(* IEC 61131-3 sources: Lasal-MCP/examples/SampleSource/2_PumpControlSolution/Stations/MachineControl/MachineControl/Class/SafetyCDIAS_Base (part 2) *)

        p_HandlePDOWrite^$USINT := VARAN_DO_NO_RUN;
      end_if;

      ud_LocalMoveDestAddr := pPDOWriteData$UDINT;
    end_if;

    if sd_VaranType = 1 then

      //add data object for TDO write
      sd_retval := MasterConnect.AddWrDO( ud_dol_type   := VARAN_DOL_ISO
                                        , p_ud_handle	  := ( #p_HandleTDOWrite )$^UDINT
                                        , ud_address	  := ui_MyPlace + OFFSET_STDO_DATA
                                        , ud_length	    := STDO_LENGTH
                                        , p_ud_data	    := ( #p_us_Handle_TDO_Write )$^UDINT
                                        , ud_type			  := 1
                                        );

      //look for an error
      if ( sd_retval <> 0 ) then
        State.uiIO_Flags				          := 0;
        State.uiIO_Flags.NoCalibration	  := 1;
        State.uiIO_Flags.PhysicAccessOff  := 1;
        return;
      end_if;
    else  // for mover we have to say it's a single execution

      //add data object for TDO write
      sd_retval := MasterConnect.AddWrDO( ud_dol_type   := VARAN_DOL_ISO
                                        , p_ud_handle	  := ( #p_HandleTDOWrite )$^UDINT
                                        , ud_address	  := ui_MyPlace + OFFSET_STDO_DATA
                                        , ud_length	    := STDO_LENGTH
                                        , p_ud_data	    := ( #p_us_Handle_TDO_Write )$^UDINT
                                        , ud_type			  := 1 OR VM_SINGLE_ID
                                        );

      //look for an error
      if ( sd_retval <> 0 ) then
        State.uiIO_Flags				          := 0;
        State.uiIO_Flags.NoCalibration	  := 1;
        State.uiIO_Flags.PhysicAccessOff  := 1;
        return;
      end_if;

      (p_HandleTDOWrite$^USINT )^ := VARAN_DO_NO_RUN;
    end_if;

    // only for modules with outputs
    if Kennung <> CSDI16x_ID then

      //add data object for unsafe output write
      sd_retval := MasterConnect.AddWrDO( ud_dol_type   := VARAN_DOL_ISO
                                        , p_ud_handle	  := ( #p_HandleUnsafeOutWrite )$^UDINT
                                        , ud_address	  := ui_MyPlace + OFFSET_UNSAFE_VAR
                                        , ud_length	    := UNSAFE_OUT_LENGTH
                                        , p_ud_data	    := ( #p_ui_UnsafeOutWrite )$^UDINT
                                        , ud_type			  := 1
                                        );

      //look for an error
      if ( sd_retval <> 0 ) then
        State.uiIO_Flags				          := 0;
        State.uiIO_Flags.NoCalibration	  := 1;
        State.uiIO_Flags.PhysicAccessOff  := 1;
        return;
      end_if;
    end_if;

    //data object for LEDs, SSDO State, STDO State, SPDO DataLength and time sync handshake
    sd_retval := MasterConnect.AddRdDO( ud_dol_type   := VARAN_DOL_ISO
                                      , p_ud_handle   := ( #p_HandleLED )$^UDINT
                                      , ud_address    := ui_MyPlace + OFFSET_LED
                                      , ud_length     := 15
                                      , p_ud_data     := ( #p_ud_Handle_LED )$^UDINT
                                      , ud_type       := 1
                                      );

    //look for an error
    if ( sd_retval <> 0 ) then
      State.uiIO_Flags				          := 0;
      State.uiIO_Flags.NoCalibration	  := 1;
      State.uiIO_Flags.PhysicAccessOff  := 1;
      return;
    end_if;

    p_us_Handle_TDO_Read_Length   := p_ud_Handle_LED + (OFFSET_STDO_STATUS - OFFSET_LED);
    p_us_Handle_TDO_Read_Length^  := 0;

    pPDOReadLengthData := p_ud_Handle_LED + (OFFSET_SPDO_LENGTH - OFFSET_LED);
    pPDOReadLengthData^ := 0;

    p_us_Handle_TDO_Status_Write  := p_ud_Handle_LED + (OFFSET_STDO_STATUS_WRITE - OFFSET_LED);
    p_us_Handle_TDO_Status_Write^ := 0;

    p_us_Handle_TimeSyncHS_Read   := p_ud_Handle_LED + (OFFSET_TIMESYNC_HANDSHAKE - OFFSET_LED);
    p_us_Handle_TimeSyncHS_Read^  := 0;

    if sd_VaranType = 1 then

      //add data object for time sync handshake
      sd_retval := MasterConnect.AddWrDO( ud_dol_type   := VARAN_DOL_ISO
                                        , p_ud_handle	  := ( #p_Handle_TimeSyncHS_Write )$^UDINT
                                        , ud_address	  := ui_MyPlace + OFFSET_TIMESYNC_HANDSHAKE
                                        , ud_length	    := 1
                                        , p_ud_data	    := ( #p_us_Handle_TimeSyncHS_Write )$^UDINT
                                        , ud_type			  := 1
                                        );

    else  // for mover we have to say it's a single execution

      //add data object for TDO write
      sd_retval := MasterConnect.AddWrDO( ud_dol_type   := VARAN_DOL_ISO
                                        , p_ud_handle	  := ( #p_Handle_TimeSyncHS_Write )$^UDINT
                                        , ud_address	  := ui_MyPlace + OFFSET_TIMESYNC_HANDSHAKE
                                        , ud_length	    := 1
                                        , p_ud_data	    := ( #p_us_Handle_TimeSyncHS_Write )$^UDINT
                                        , ud_type			  := 1 OR VM_SINGLE_ID
                                        );
      (p_Handle_TimeSyncHS_Write$^USINT )^ := VARAN_DO_NO_RUN;
    end_if;

    //look for an error
    if ( sd_retval <> 0 ) then
      State.uiIO_Flags				          := 0;
      State.uiIO_Flags.NoCalibration	  := 1;
      State.uiIO_Flags.PhysicAccessOff  := 1;
      return;
    end_if;

    //add data object for TDO read
    sd_retval := MasterConnect.AddRdDO( ud_dol_type   := VARAN_DOL_ISO
                                      , p_ud_handle	  := ( #p_HandleTDORead )$^UDINT
                                      , ud_address	  := ui_MyPlace + OFFSET_STDO_DATA
                                      , ud_length	    := STDO_LENGTH
                                      , p_ud_data	    := ( #p_us_Handle_TDO_Read )$^UDINT
                                      , ud_type			  := 1
                                      );

    //look for an error
    if ( sd_retval <> 0 ) then
      State.uiIO_Flags				          := 0;
      State.uiIO_Flags.NoCalibration	  := 1;
      State.uiIO_Flags.PhysicAccessOff  := 1;
      return;
    end_if;

    // fast unsafe variables (only if activated)
    if ActivateFastUnsafeIOs then
      //add data object for fast unsafe output and input variables
      sd_retval :=  MasterConnect.AddRdWrDO(ud_dol_type       := VARAN_DOL_ISO
                                          , p_ud_handle       := ( #p_HandleFastUnsafeIOs )$^UDINT
                                          , ud_address_read   := ui_MyPlace + OFFSET_FAST_UNSAFE_IOS
                                          , ud_length_read    := 1
                                          , p_ud_data_read    := ( #p_us_Handle_FastUnsafeOutputs )$^UDINT
                                          , ud_address_write  := ui_MyPlace + OFFSET_FAST_UNSAFE_IOS
                                          , ud_length_write   := 1
                                          , p_ud_data_write   := ( #p_us_Handle_FastUnsafeInputs )$^UDINT
                                          , ud_type           := 1
                                          );

      //look for an error
      if ( sd_retval <> 0 ) then
        State.uiIO_Flags				          := 0;
        State.uiIO_Flags.NoCalibration	  := 1;
        State.uiIO_Flags.PhysicAccessOff  := 1;
        return;
      end_if;
    end_if;
  end_if;

END_FUNCTION

FUNCTION VIRTUAL SafetyCDIAS_Base::GetPointer2PDOBuffer
	VAR_OUTPUT
		ud_PDOBuffer 	: UDINT;
	END_VAR

  PDOOutputIsUsed := TRUE;

  //set pointer to address of buffer pointer
  ud_PDOBuffer := ( #PDOOutputBuffer )$UDINT;

END_FUNCTION

FUNCTION VIRTUAL SafetyCDIAS_Base::AddRoutingElement
	VAR_INPUT
		ud_SafeNumber 	: HDINT;
		ud_thisp 	      : UDINT;
		pObject 	      : ^PathInfoType;
	END_VAR
	VAR_OUTPUT
		sd_retval 	    : DINT;
	END_VAR
  VAR
  	p_RoutElement   : ^RoutElement;
    ui_PathLength   : UINT;
    NewElement      : BOOL;
  END_VAR

  if ( ( ud_SafeNumber <> 0 ) & ( ud_thisp <> NIL ) ) then
    if ui_CntRoutElements < MAX_NUMBER_ROUT_ELEMENTS then

      NewElement := TRUE;

      if ui_CntRoutElements then
        //check if object this-pointer already exists in routing table
        p_RoutElement := GetRoutingElementByThis( ud_thisp := ud_thisp );
      else
        p_RoutElement := NIL;
      end_if;

      if p_RoutElement = NIL then
        //add new element

        //set pointer to empty element on last position
        p_RoutElement := p_RoutTable + ( ui_CntRoutElements ) * sizeof(RoutElement);
      else
        // we don't have a new element, we just update an existing
        NewElement := FALSE;
      end_if;

      //add path

      // path isn't stored if it's the routing table of safe input module, because
      // it doesn't need the information
      if pObject^.p_us_Path & pObject^.p_us_PathComp
         & ((NewElement = TRUE) | ((NewElement = FALSE) & (p_RoutElement^.p_CompressedPath = NIL) & (p_RoutElement^.ui_ComprPathLen = 0))) // only if it isn't already set
         then

        // the whole object path isn't stored, because the path can't be used for routing of SDOs;
        // The length of the path varies and it's possible, that the path is too long
        // to transfer it in SDO header. Instead of it the compressed path is used for addressing.

        ui_PathLength := pObject^.ui_PathCompLen;
        p_RoutElement^.p_CompressedPath$pVoid := To_StdLib.Malloc(size := ui_PathLength);

        if ( p_RoutElement^.p_CompressedPath = NIL ) then

          State.uiIO_Flags                  := 0;
          State.uiIO_Flags.PhysicAccessOff 	:= 1;
          sd_retval                         :=-1;
          ClassState := _MemAllocFailed;
          return;

        end_if;

        // store compressed path into actual routing element
        To_StdLib.MemCpy(dest := p_RoutElement^.p_CompressedPath, source := pObject^.p_us_PathComp, size := ui_PathLength);
        p_RoutElement^.ui_ComprPathLen := ui_PathLength;
      elsif NewElement then

        // not routing table of safety CPU of safety output
        p_RoutElement^.p_CompressedPath := NIL;
        p_RoutElement^.ui_ComprPathLen  := 0;
      end_if;

      //insert data
      p_RoutElement^.ud_SafeNumber      := ud_SafeNumber;
      p_RoutElement^.ud_thisp           := ud_thisp;

      if NewElement then
        //increase counter
        ui_CntRoutElements += 1;
      end_if;

      sd_retval := 0;
    else

      sd_retval := -1;
      LogError("@ZZZZ (SafetyCDIAS_Base::AddRoutingElement) Maximum number of possible routing elements reached");
    end_if;
  else

    sd_retval := -1;

    if ud_SafeNumber = 0 then
      LogError("@ZZZZ (SafetyCDIAS_Base::AddRoutingElement) 0 is an invalid safety number");
    else
      LogError("@ZZZZ (SafetyCDIAS_Base::AddRoutingElement) NIL pointer given as this pointer");
    end_if;
  end_if;

END_FUNCTION

FUNCTION VIRTUAL SafetyCDIAS_Base::GetRoutingPointerByNumber
	VAR_INPUT
		ud_SafeNumber 	: HDINT;
	END_VAR
	VAR_OUTPUT
		ud_thisp 	      : UDINT;
	END_VAR
  VAR
  	i               : UINT;
    p_RoutElement   : ^RoutElement;
  END_VAR

  ud_thisp := 0;

  //no valid safety number
  if ( ud_SafeNumber = 0 ) then
    return;
  end_if;

  //set pointer on first routing element
  p_RoutElement := p_RoutTable;

  //check each element
  if ( ui_CntRoutElements > 0 ) then
    for i := 0 to ui_CntRoutElements - 1 by 1 do

      //if searched safety number is found, this-pointer is returned
      if ( p_RoutElement^.ud_SafeNumber = ud_SafeNumber ) then

        ud_thisp := p_RoutElement^.ud_thisp;
        return;

      end_if;

      //set pointer to next element
      p_RoutElement += sizeof ( RoutElement );

    end_for;
  end_if;

END_FUNCTION

FUNCTION VIRTUAL SafetyCDIAS_Base::GetRoutingPointerByPath
	VAR_INPUT
		p_ActObjectPath 	: ^USINT;
		ActPathLen 	      : UINT;
	END_VAR
	VAR_OUTPUT
		ud_thisp          : UDINT;
	END_VAR
  VAR
  	i                 : UINT;
    p_RoutElement     : ^RoutElement;
    retcode           : UINT;
  END_VAR

  ud_thisp := 0;

  //set pointer on first routing element
  p_RoutElement := p_RoutTable;

  //check each element
  if ( ui_CntRoutElements > 0 ) then
    for i := 0 to ui_CntRoutElements - 1 by 1 do

      if p_RoutElement^.p_CompressedPath & (p_RoutElement^.ui_ComprPathLen = ActPathLen) then

        //if searched path is found, this-pointer is returned
        retcode := To_StdLib.MemCmp(dest:= p_ActObjectPath, source:= p_RoutElement^.p_CompressedPath , size:= ActPathLen);

        if retcode = 0 then

          ud_thisp := p_RoutElement^.ud_thisp;
          return;

        end_if;
      end_if;

      //set pointer to next element
      p_RoutElement += sizeof ( RoutElement );

    end_for;
  end_if;

END_FUNCTION

FUNCTION VIRTUAL SafetyCDIAS_Base::ConfigSafetyInput
	VAR_INPUT
		ud_SafeNrCPU 	        : HDINT;
		ud_thisp 	            : UDINT;
		p_PDOBuffer 	        : ^UDINT;
		pMoveActive 	        : ^PDOMoveState;
		p_ud_HandleSourceDO 	: ^UDINT;
		p_ud_MoveSourceAddr 	: ^UDINT;
		p_ud_MoveSourceOffset : ^UDINT;
	END_VAR
	VAR_OUTPUT
		ud_SafeNrModul 	      : HDINT;
	END_VAR
  VAR
  	TempPathInfo          : PathInfoType;
  END_VAR

  ud_SafeNrModul := 0;

  if (State.uiIO_Flags = 0) then
    if ( ud_SafeNrCPU ) then

      // if pMoveActive is available, the data are sent to a CPU via VARAN => moving is possible
      if pMoveActive then
        // if input module is also accessed via VARAN => activate moving
        if b_VaranAvailable & (b_SafetyOnLocalCDIAS = FALSE) then
          // pdos are moved from csdi to cscp
          b_MoveCommandOutputActive := _Active;

          p_ud_MoveSourceAddr^      := pPDOReadData$UDINT;

          // Return DO Handle and Offset, Needed for Payload Move DOs
          if sd_VaranType = 1 then  // Return DO Handle
            p_ud_HandleSourceDO^    := p_HandlePDORead$UDINT;
          else                      // Return VaranDataMoversDO Handle
            p_ud_HandleSourceDO^    := 0;
          end_if;

          p_ud_MoveSourceOffset^    := 0;

          // Return DO Handle and Offset, Needed for Payload Move DOs
          if sd_VaranType = 1 then  // Return DO Handle
            p_ud_HandleSourceDO^    := p_HandlePDORead$UDINT;
          else                      // Return VaranDataMoversDO Handle
            p_ud_HandleSourceDO^    := ud_HandlePDOReadMoverDO;
          end_if;

          p_ud_MoveSourceOffset^    := 0;
        else
          // pdos are not moved from csdi to cscp or cscp to csto
          pMoveActive^              := _Inactive;
          b_MoveCommandOutputActive := _Inactive;
        end_if;
      else
        b_MoveCommandOutputActive   := _Inactive;
      end_if;

      // we start the data object for continous writing to the module after we know that there is an input for this module and the move command is active
      if b_VaranAvailable & (b_MoveCommandOutputActive = _Active) then
        if sd_VaranType = 1 then
          if StartRtDOs = 0 then
            StartRtDOs := 1;
          end_if;
        end_if;
      end_if;

      InitPathInfo(#TempPathInfo);

      //add CPU to routing table for SDO
      if ( AddRoutingElement( ud_SafeNumber   := ud_SafeNrCPU
                            , ud_thisp        := ud_thisp
                            , pObject         := #TempPathInfo
                            ) = 0 ) then

        //return own safety number
        ud_SafeNrModul := SafetyNumber;

      end_if;

      //set pointer to address of buffer pointer
      p_PDOBuffer^ := GetPointer2PDOBuffer();
    else
      LogError("@ZZZZ (SafetyCDIAS_Base::ConfigSafetyInput) 0 is an invalid safety number for the safety CPU");
      b_ReInitMarker := TRUE;
    end_if;
  else
    LogError("@ZZZZ (SafetyCDIAS_Base::ConfigSafetyInput) A module with safety outputs, which is used in the safety CPU configuration is not available");
    b_ReInitMarker := TRUE;
  end_if;

END_FUNCTION

FUNCTION VIRTUAL SafetyCDIAS_Base::ConfigSafetyOutput
	VAR_INPUT
		ud_SafeNrCPU 	      : HDINT;
		ud_thisp 	          : UDINT;
		ud_p_PDOBuffer 	    : UDINT;
		pObject 	          : ^PathInfoType;
		pMoveActive 	      : ^PDOMoveState;
    ud_HandleSourceDO   : UDINT;
		ud_MoveSourceAddr   : UDINT;
    ud_MoveSourceOffset : UDINT;
    b_IsOptional        : BOOL;
	END_VAR
	VAR_OUTPUT
		ud_SafeNrModul      : HDINT;
	END_VAR
  VAR
  	i                   : DINT;
  END_VAR

  ud_SafeNrModul := 0;

  if (State.uiIO_Flags = 0) then
    if ( ud_SafeNrCPU ) then

      //add CPU to routing table for SDO
      if ( AddRoutingElement( ud_SafeNumber   := ud_SafeNrCPU
                            , ud_thisp        := ud_thisp
                            , pObject         := pObject
                            ) = 0 ) then

        //return own safety number and object path
        ud_SafeNrModul := SafetyNumber;

      end_if;

      //add PDO of CPU to list of input elements
      AddPDOToInputBuffer(ud_p2Buffer         := ud_p_PDOBuffer
                        , ud_HandleSourceDO   := ud_HandleSourceDO
                        , ud_MoveSourceAddr   := ud_MoveSourceAddr
                        , ud_MoveSourceOffset :=ud_MoveSourceOffset
                        , ud_SafetyNr         := ud_SafeNrCPU
                        , b_IsOptional        := b_IsOptional
                        );

      // if we got an adress of the source data from cpu, the cpu must be connected via VARAN => moving is possible
      if ud_MoveSourceAddr then

        // if output module is also accessed via VARAN => activate moving
        if b_VaranAvailable & (b_SafetyOnLocalCDIAS = FALSE) then
          // pdos are moved from cscp to csto
          b_MoveCommandInputActive  := _Active;
        else
          // pdos are not moved from cscp to csto because csto is not connected via VARAN
          if pMoveActive then
            pMoveActive^            := _Inactive;
          end_if;
          b_MoveCommandInputActive  := _Inactive;
        end_if;
      else
        // pdos are not moved from cscp to csto because cscp (and/or csto) is not connected via VARAN
        if pMoveActive then
          pMoveActive^              := _Inactive;
        end_if;
        b_MoveCommandInputActive    := _Inactive;
      end_if;

      // we start the data object for continous writing to the module after we know that there is an input for this module and the move command is active
      if b_VaranAvailable & (b_MoveCommandInputActive = _Active) then
        b_StartDOs := TRUE;
      elsif b_VaranAvailable & (sd_VaranType = 1) then
        MasterConnect.ResetDO( p_data_object := p_HandlePDOWrite$^DINT, us_state := VARAN_DO_NO_RUN, ud_bytes := MaxLengthPDOWrite);

        if AdditionalSPDOs & (ui_cnt_PDOInputBuffer > 1) then
          if AdditionalSPDOs > (ui_cnt_PDOInputBuffer-1) then
            AdditionalSPDOs := ui_cnt_PDOInputBuffer-1;
          end_if;

          for i := 0 to (AdditionalSPDOs-1) do
            MasterConnect.ResetDO( p_data_object := aAdditionalPDOs[i].p_HandlePDOWrite$^DINT, us_state := VARAN_DO_NO_RUN, ud_bytes := MaxLengthPDOWrite);
          end_for;
        end_if;
      end_if;
    else
      LogError("@ZZZZ (SafetyCDIAS_Base::ConfigSafetyOutput) 0 is an invalid safety number for the safety CPU");
      b_ReInitMarker := TRUE;
    end_if;
  else
    LogError("@ZZZZ (SafetyCDIAS_Base::ConfigSafetyOutput) A module with safety outputs, which is used in the safety CPU configuration is not available");
    b_ReInitMarker := TRUE;
  end_if;

END_FUNCTION

FUNCTION VIRTUAL SafetyCDIAS_Base::ConfigSafetyCPU
	VAR_OUTPUT
		ud_SafeNrModul 	: HDINT;
	END_VAR

  //return own safety number
  ud_SafeNrModul := SafetyNumber;

END_FUNCTION

FUNCTION VIRTUAL SafetyCDIAS_Base::AddPDOToInputBuffer
	VAR_INPUT
		ud_p2Buffer 	        : UDINT;
		ud_HandleSourceDO 	  : UDINT;
		ud_MoveSourceAddr 	  : UDINT;
		ud_MoveSourceOffset 	: UDINT;
		ud_SafetyNr 	        : HDINT;
		b_IsOptional 	        : BOOL;
		us_PdoLen 	          : USINT;
	END_VAR
	VAR_OUTPUT
		sd_retval 	          : DINT;
	END_VAR
  VAR
  	p_BufferElement       : ^PDOInputBuffer;
  END_VAR

  sd_retval := 0;

  //check if input buffer is already in list
  p_BufferElement := GetPDOInputBuffer(ud_p2Buffer := ud_p2Buffer);

  //buffer already in list -> do nothing
  if ( p_BufferElement ) then
    return;
  else
    aPDOInputBuffer[ui_cnt_PDOInputBuffer].ud_p2Buffer        := ud_p2Buffer;
    aPDOInputBuffer[ui_cnt_PDOInputBuffer].ud_HandleSourceDO  := ud_HandleSourceDO;   //LanSte 28.05.2013 For Payload support
    aPDOInputBuffer[ui_cnt_PDOInputBuffer].ud_MoveSourceAddr  := ud_MoveSourceAddr;
    aPDOInputBuffer[ui_cnt_PDOInputBuffer].ud_MoveSourceOffset:= ud_MoveSourceOffset; //LanSte 28.05.2013 For Payload support
    //*****************************************************************************

    aPDOInputBuffer[ui_cnt_PDOInputBuffer].b_TimeSynchron     := FALSE;
    aPDOInputBuffer[ui_cnt_PDOInputBuffer].ud_SafetyNr        := ud_SafetyNr;
    aPDOInputBuffer[ui_cnt_PDOInputBuffer].us_PDOLen          := us_PDOLen;
    aPDOInputBuffer[ui_cnt_PDOInputBuffer].b_IsOptional       := b_IsOptional;

    if ui_cnt_PDOInputBuffer = 0 then
      // only when adding the first input PDO we increment our module counter
      ModuleSyncNo += 1;
    end_if;

    ui_cnt_PDOInputBuffer += 1;
  end_if;

END_FUNCTION

FUNCTION VIRTUAL SafetyCDIAS_Base::WritePDO2Module
  VAR
    p_PDOInBufferAct  : ^PDOInputBuffer;
    p_PDO_data        : ^UINT;
    PDOLength         : USINT;
    p_addressWr		    : ^VaranDOSettingsWr;
    i                 : DINT;
  END_VAR

  // if last PDO was selected (or a PDO which doesn't exist anymore), select first
  if ( ui_cnt_PDOInBufferAct >= ui_cnt_PDOInputBuffer ) then
    ui_cnt_PDOInBufferAct := 0;
  end_if;

  p_PDOInBufferAct := #aPDOInputBuffer[ui_cnt_PDOInBufferAct];

  if b_MoveCommandInputActive <> _Active then
    p_PDO_data := p_PDOInBufferAct^.ud_p2Buffer$^UINT;

    // get length out of PDO frame
    PDOLength := (p_PDO_data$^USINT + PDOType.Length)^ + sizeof(PDOType.CRC);

    //Save length to variable
    PDOWriteLen := PDOLength;

    // only if length is bigger than minimum and smaller than maximum
    if ( PDOLength > PDOType.Length ) & ( PDOLength <= SPDO_MAX_LENGTH ) then
  #ifdef SAFETY_OVER_DIAS
      if ( b_im ) then

        //copy word by word
        for i := 0 to ((PDOLength/2)-1) by 1 do

          (( a_Handle_PDO_Write[i] )$^UINT )^ := ( p_PDO_data + ( i * 2 ))^;

        end_for;

      else
  #endif

        //copy whole PDO
        To_StdLib.MemCpy(dest := pPDOWriteData, source := p_PDO_data, size := PDOLength);

#ifdef DO_DEBUG
        DOCheck(pFrame:=p_PDO_data$^SDOStdHeader, pCheckStruct:=#PDOWrite);
#endif

#ifdef SAFETY_PROTOCOL_ANALYZER_ACTIVATED
  RecordFrame(p_PDO_data$^DINT, 1);
#endif

        if b_VaranAvailable then

          if b_PayloadSupport then

            if (sd_VaranType = 1) then

            // correct size of data object to PDOLength
              ChangeDOLengthOffset( ud_DOHandle     := p_HandlePDOWrite$UDINT
                                  , ud_length_write := PDOLength
                                  );
              EnableDO(ud_DOHandle := p_HandlePDOWrite$UDINT );
              PDOSingleRunActive := 2;  // No singlerun with Payload
            else
              p_HandlePDOWriteEnable^ := VARAN_MOVER_DO_CONT_RUN;
              PDOSingleRunActive := 2;
            end_if;

          else
            if (sd_VaranType = 1) then

              // correct size of data object to PDOLength
              p_addressWr := pPDOWriteData - sizeof(VaranDOSettingsWr);
              p_addressWr^.us_ByteCnt := PDOLength;
              p_HandlePDOWrite^.usSendBufferLength := sizeof(VaranDOSettingsWr) + to_uint(PDOLength);

              p_HandlePDOWrite^.ucCtrlStat := VARAN_DO_SINGLE_RUN;
            else
              (p_HandlePDOWrite$^USINT )^ := VARAN_MOVER_DO_CONT_RUN;
              PDOSingleRunActive := 2;  // This Marker is also used for aAdditionalPDOs
            end_if;

          end_if;

        end_if;

        if AdditionalSPDOs then

          for i := 0 to (AdditionalSPDOs-1) do

            //increase counter for pointer position for next PDO
            ui_cnt_PDOInBufferAct += 1;

            //if last PDO was read, reset counter for first PDO
            if ( ui_cnt_PDOInBufferAct = ui_cnt_PDOInputBuffer ) then
              ui_cnt_PDOInBufferAct := 0;
            end_if;

            p_PDOInBufferAct := #aPDOInputBuffer[ui_cnt_PDOInBufferAct];

            p_PDO_data := p_PDOInBufferAct^.ud_p2Buffer$^UINT;

            // get length out of PDO frame
            PDOLength := (p_PDO_data$^USINT + PDOType.Length)^ + sizeof(PDOType.CRC);

            // only if length is bigger than minimum and smaller than maximum
            if ( PDOLength > PDOType.Length ) & ( PDOLength <= SPDO_MAX_LENGTH ) then

              //copy whole PDO
              To_StdLib.MemCpy(dest := aAdditionalPDOs[i].pPDOWriteData, source := p_PDO_data, size := PDOLength);

#ifdef DO_DEBUG
              DOCheck(pFrame:=p_PDO_data$^SDOStdHeader, pCheckStruct:=#PDOWrite);
#endif

#ifdef SAFETY_PROTOCOL_ANALYZER_ACTIVATED
  RecordFrame(p_PDO_data$^DINT, 1);
#endif

              if b_VaranAvailable then
                if b_PayloadSupport then
                  if (sd_VaranType = 1) then
                  // correct size of data object to PDOLength
                    ChangeDOLengthOffset( ud_DOHandle     := aAdditionalPDOs[i].p_HandlePDOWrite$UDINT
                                        , ud_length_write := PDOLength
                                        );
                    EnableDO(ud_DOHandle := aAdditionalPDOs[i].p_HandlePDOWrite$UDINT); // PDOSingleRunActive is used to deactivates these again

                  else
                    aAdditionalPDOs[i].p_HandlePDOWriteEnable^ := VARAN_MOVER_DO_CONT_RUN;  // PDOSingleRunActive is used to deactivates these again
                  end_if;
                else
                  if (sd_VaranType = 1) then
                      // correct size of data object to PDOLength
                    p_addressWr := aAdditionalPDOs[i].pPDOWriteData - sizeof(VaranDOSettingsWr);
                    p_addressWr^.us_ByteCnt := PDOLength;
                    aAdditionalPDOs[i].p_HandlePDOWrite^.usSendBufferLength := sizeof(VaranDOSettingsWr) + to_uint(PDOLength);

                    aAdditionalPDOs[i].p_HandlePDOWrite^.ucCtrlStat := VARAN_DO_SINGLE_RUN;
                  else
                    (aAdditionalPDOs[i].p_HandlePDOWrite$^USINT )^ := VARAN_MOVER_DO_CONT_RUN;  // PDOSingleRunActive is used to deactivates these again
                  end_if;
                end_if;
              end_if;
            end_if;
          end_for;
        end_if;
  #ifdef SAFETY_OVER_DIAS
      end_if;
  #endif
    end_if;
  else
    if (p_PDOInBufferAct^.ud_MoveSourceAddr) then

#ifdef VM_DEBUG_PAYLOAD
      if b_PayloadSupport = true &
        p_PDOInBufferAct^.ud_HandleSourceDO = 0 then
        // Handle mus be valid with payload support
        ((0)$^USINT)^ := 0;
      end_if;
#endif

      PDOLength := ((p_PDOInBufferAct^.ud_MoveSourceAddr)$^USINT + PDOType.Length)^ + sizeof(PDOType.CRC);

      //Save length to variable
      PDOWriteLen := PDOLength;

      if ( PDOLength > PDOType.Length ) & ( PDOLength <= MaxLengthPDOWrite) then

        if (sd_VaranType = 1) then

          if b_PayloadSupport then
          // correct size of data object to PDOLength
            ChangeDOLengthOffset( ud_DOHandle     := p_HandlePDOWrite$UDINT
                                , ud_length_write := PDOLength
                                );
            //start data object
            EnableDO(ud_DOHandle := p_HandlePDOWrite$UDINT);
          else
            // correct size of data object to PDOLength
            p_addressWr := pPDOWriteData - sizeof(VaranDOSettingsWr);
            p_addressWr^.us_ByteCnt := PDOLength;
            p_HandlePDOWrite^.usSendBufferLength := sizeof(VaranDOSettingsWr) + to_uint(PDOLength);

            //start data object
            MasterConnect.ResetDO( p_data_object := p_HandlePDOWrite$^DINT, us_state := VARAN_DO_CONT_RUN, ud_bytes := PDOLength );
          end_if;

        elsif b_PayloadSupport = false then // No Payload + Mover
          PDOLength := MaxLengthPDOWrite-1;
        end_if;

        if b_PayloadSupport then

          if sd_VaranType = 1 then
            ChangeMovDOLengthOffset(ud_MovDOHandle              := InputMovHandle$UDINT
                                  , ud_sourceReadDOHandle       := p_PDOInBufferAct^.ud_HandleSourceDO
                                  , ud_SourceReadOffset         := p_PDOInBufferAct^.ud_MoveSourceOffset
                                  , ud_destinationWriteDOHandle := p_HandlePDOWrite$UDINT
                                  , ud_DestinationWriteOffset   := 0
                                  , ud_lengthmove               := PDOLength);
          else  // VaranDatamover
            ChangeMovDOLengthOffset(ud_MovDOHandle              := InputMovHandle$UDINT
                                  , ud_sourceReadDOHandle       := p_PDOInBufferAct^.ud_HandleSourceDO
                                  , ud_SourceReadOffset         := p_PDOInBufferAct^.ud_MoveSourceOffset
                                  , ud_destinationWriteDOHandle := ud_HandlePDOWriteMoverDO
                                  , ud_DestinationWriteOffset   := 0
                                  , ud_lengthmove               := PDOLength);
          end_if;

          // moving is done every cycle
          EnableDO(ud_DOHandle := InputMovHandle$UDINT);

        else
          InputMovSettings^.ud_AddressDest := ud_LocalMoveDestAddr;
          InputMovSettings^.ud_AddressSrc  := p_PDOInBufferAct^.ud_MoveSourceAddr;
          InputMovSettings^.ui_ByteCnt     := PDOLength;

          // moving is done every cycle
          InputMovHandle^.ucCtrlStat := VARAN_DO_CONT_RUN;
        end_if;

        if AdditionalSPDOs then

          for i := 0 to (AdditionalSPDOs-1) do

            //increase counter for pointer position for next PDO
            ui_cnt_PDOInBufferAct += 1;

            //if last PDO was read, reset counter for first PDO
            if ( ui_cnt_PDOInBufferAct = ui_cnt_PDOInputBuffer ) then
              ui_cnt_PDOInBufferAct := 0;
            end_if;

            p_PDOInBufferAct := #aPDOInputBuffer[ui_cnt_PDOInBufferAct];

            if p_PDOInBufferAct^.ud_MoveSourceAddr then
              PDOLength := ((p_PDOInBufferAct^.ud_MoveSourceAddr)$^USINT + PDOType.Length)^ + sizeof(PDOType.CRC);

              if ( PDOLength > PDOType.Length ) & ( PDOLength <= MaxLengthPDOWrite) then

                if (sd_VaranType = 1) then

                  if b_PayloadSupport then

                  // correct size of data object to PDOLength
                    ChangeDOLengthOffset( ud_DOHandle     := aAdditionalPDOs[i].p_HandlePDOWrite$UDINT
                                        , ud_length_write := PDOLength
                                        );

                    //start data object
                    EnableDO(ud_DOHandle := aAdditionalPDOs[i].p_HandlePDOWrite$UDINT);
                  else
                    // correct size of data object to PDOLength
                    p_addressWr := aAdditionalPDOs[i].pPDOWriteData - sizeof(VaranDOSettingsWr);
                    p_addressWr^.us_ByteCnt := PDOLength;
                    aAdditionalPDOs[i].p_HandlePDOWrite^.usSendBufferLength := sizeof(VaranDOSettingsWr) + to_uint(PDOLength);

                    //start data object
                    MasterConnect.ResetDO( p_data_object := aAdditionalPDOs[i].p_HandlePDOWrite$^DINT, us_state := VARAN_DO_CONT_RUN, ud_bytes := PDOLength );
                  end_if;

                elsif b_PayloadSupport = false then // No Payload Mover
                  PDOLength := MaxLengthPDOWrite-1;
                end_if;
              end_if;

              if b_PayloadSupport then
                if sd_VaranType = 1 then
                  ChangeMovDOLengthOffset(ud_MovDOHandle              := aAdditionalPDOs[i].InputMovHandle$UDINT
                                        , ud_sourceReadDOHandle       := p_PDOInBufferAct^.ud_HandleSourceDO
                                        , ud_SourceReadOffset         := p_PDOInBufferAct^.ud_MoveSourceOffset
                                        , ud_destinationWriteDOHandle := aAdditionalPDOs[i].p_HandlePDOWrite$UDINT
                                        , ud_DestinationWriteOffset   := 0
                                        , ud_lengthmove               := PDOLength);
                else  // VaranDataMover
                  ChangeMovDOLengthOffset(ud_MovDOHandle              := aAdditionalPDOs[i].InputMovHandle$UDINT
                                        , ud_sourceReadDOHandle       := p_PDOInBufferAct^.ud_HandleSourceDO
                                        , ud_SourceReadOffset         := p_PDOInBufferAct^.ud_MoveSourceOffset
                                        , ud_destinationWriteDOHandle := aAdditionalPDOs[i].ud_HandlePDOWriteMoverDO
                                        , ud_DestinationWriteOffset   := 0
                                        , ud_lengthmove               := PDOLength);
                end_if;
                // moving is done every cycle
                EnableDO(ud_DOHandle := aAdditionalPDOs[i].InputMovHandle$UDINT);
              else
                aAdditionalPDOs[i].InputMovSettings^.ud_AddressDest := aAdditionalPDOs[i].ud_LocalMoveDestAddr;
                aAdditionalPDOs[i].InputMovSettings^.ud_AddressSrc  := p_PDOInBufferAct^.ud_MoveSourceAddr;
                aAdditionalPDOs[i].InputMovSettings^.ui_ByteCnt     := PDOLength;

                // moving is done every cycle
                aAdditionalPDOs[i].InputMovHandle^.ucCtrlStat       := VARAN_DO_CONT_RUN;
              end_if;

            end_if;
          end_for;
        end_if;
      end_if;
    else
      bd_LogOnceMarker.MoveSourceInvalid := TRUE;
    end_if;
  end_if;

  //increase counter for pointer position for next PDO
  ui_cnt_PDOInBufferAct += 1;

  //if last PDO was read, reset counter for first PDO
  if ( ui_cnt_PDOInBufferAct = ui_cnt_PDOInputBuffer ) then
    ui_cnt_PDOInBufferAct := 0;
  end_if;

END_FUNCTION

FUNCTION VIRTUAL SafetyCDIAS_Base::Varan_CallbackSafe
	VAR_INPUT
		ud_reason 	: UDINT;
	END_VAR
  VAR
		MyPara 	    : CmdStruct;
		MyResult	  : results;
  END_VAR

	//look for reason
	if ( ud_reason = 0 ) then		//connect
    if b_PayloadSupport & (sd_VaranType = 2) then
      if ( AddDO() ) then

        return;

      end_if;
    end_if;
		//read Kennung
		Kennung := MasterConnect.GetKennung( Place );

    // Only Read Serial No if Kennung was successfully read. Otherwise we get an EPROM Error at the CIV even if the module is not required
    if Kennung & Kennung <> 16#ff then
      GetSerialNo();
    end_if;

		//check right module id
	 	if ( Kennung = ud_MyModuleID ) then

      // get variant from eeprom
      us_Variant := 16#FF;
      MasterConnect.I2CReadOneByte( AdressCDIAS := ui_MyPlace + 3
                                  , pData       := #us_Variant
                                  );

      // check variant
      if CheckVariant(us_Variant) then

        MasterConnect.RdDO(ud_address:=Place*16#100 + OFFSET_FPGA_VERSION, ud_length:=1, p_ud_data:=#FPGA_Version, ud_type:=1);

        // initialize the PLL

        // get our system time
        SystemTime_ms := (MasterConnect.GetPllTime())$USINT;

        // write it in ms to the pll period register
        MasterConnect.WrDO(ud_address:=Place*16#100 + OFFSET_PLL_CONFIG2, ud_length:=1, p_ud_data:=#SystemTime_ms, ud_type:=1);

        // check what module we got for writing the sync offset
        case Kennung of
          CSDI16x_ID: // if there are only inputs
            // sync offset to the beginning of the access on the CDIAS (with the CDIAS sync)
            ui_ActIRQSyncOffset := SYNC_OFFSET_NO_DELAY;

          CSTO08x_ID, CSCP01x_ID: // if there are also outputs
            // sync offset right after the access on the CDIAS (about half a cycle later)
            ui_ActIRQSyncOffset := SYNC_OFFSET_DELAY_OUTPUTS;
        end_case;

        // write the value to the module
        MasterConnect.WrDO(ud_address:=Place*16#100 + OFFSET_SYNC_IRQ_DELAY, ud_length:=2, p_ud_data:=#ui_ActIRQSyncOffset, ud_type:=1);
        if ( sd_VaranType = 2 & b_PayloadSupport = FALSE ) then

          if ( AddDO() ) then

            return;

          end_if;

        elsif ( sd_VaranType = 1 ) then

          StartRtDOs := 2;

          //start DOs
//          StartDO();

        end_if;

        //add module to safety communication task with SDO
        if ( AddModuleToSafetyTask() ) then
          return;
        end_if;

        //read own safety number
        if ( GetSafetyNumber() ) then
          return;
        end_if;

        // initialize of length of PDO to read
        PDOReadLen  := 0;
        PDOWriteLen := 0;

        State.uiIO_Flags := 0;

        if ClassState = _ModuleNotFound then
          if ModuleSyncNo = 0 then
            ClassState := _SafetyClassOK;
          else
            ClassState := _WaitForSynchronicity;
          end_if;
        end_if;

        // whenever the postinit has passed and we got a connect (module has been plugged in after booting the application) => get it's config
        if b_PostInitPassed = TRUE then
          // start reading the config in background (if we're in init the post-init read-out will be faster)

          ClassState            := _ReinitConfig;
          b_GetNewConfiguration := TRUE;
        end_if;

        // if we we're already connected => tell the sdias manager we're back (safetythis has to be valid if b_Reconnect is set, therefore we don't have to check it here)
        if b_Reconnect then
          MyPara.uiCmd    := CMD_SM_MODULE_RECONNECT;
          MyPara.aPara[0] := THIS$DINT;
          pSafetyManagerThis^.NewInst(#MyPara, #MyResult);
        else
            // if first connect, check for the reinit marker
            // send message to safetymanager, so all modules with the reinit marker can be reinitialized
            MyPara.uiCmd    := CMD_SM_MODULE_REINIT;
            MyPara.aPara[0] := THIS$DINT;
            pSafetyManagerThis^.NewInst(#MyPara, #MyResult);

        end_if;
      else

        State.uiIO_Flags                  := 0;
        if ( Kennung = 255 ) then
          State.uiIO_Flags.NoHW           := 1;
        else
          State.uiIO_Flags.WrongHW        := 1;
        end_if;
        State.uiIO_Flags.PhysicAccessOff  := 1;

      end_if;

    else

      State.uiIO_Flags                    := 0;
			if ( Kennung = 255 ) then
				State.uiIO_Flags.NoHW             := 1;
			else
				State.uiIO_Flags.WrongHW          := 1;
			end_if;
			State.uiIO_Flags.PhysicAccessOff    := 1;

    end_if;

	else  //disconnect

    // reset variables if it's a cpu
    if GetModuleID() = CSCP01x_ID then

      // delete request
      LastRequest := _NoOpenRequest;
      ud_AsyComRetryCounter := 0; // reset retry counter

      // remove the cpu from all classes, which use it
      ResetConfig();

      if UnsafeScheduler <> UnsafeSchedulerSetBusReady then
        us_SetBusReadyState := WaitPDOsSyncron;
        UnsafeScheduler := UnsafeSchedulerSetBusReady;
      end_if;

      MaxVarsPerReadPackage   := 0;
      ReadFramesNeeded        := 0;
      MaxVarsPerWritePackage  := 0;
      WriteFramesNeeded       := 0;
    end_if;

    if ( sd_VaranType = 1 ) then

      //stop DOs
      StopDO();

    end_if;

    // reset time sync state and tell the manager
    if pSafetyManagerThis then
      MyPara.uiCmd := CMD_SM_MODULE_DISCONNECT;
      MyPara.aPara[0] := THIS$DINT;
      pSafetyManagerThis^.NewInst(#MyPara, #MyResult);

      b_Reconnect := TRUE;
    end_if;

    b_TimeSyncActive                  := FALSE;
    TimeSyncDOActive.OwnSyncActive    := 0;

    State.uiIO_Flags					        := 0;
		State.uiIO_Flags.NoHW	 			      := 1;
		State.uiIO_Flags.PhysicAccessOff  := 1;

    ClassState := _ModuleNotFound;
  end_if;

END_FUNCTION

FUNCTION VIRTUAL GLOBAL SafetyCDIAS_Base::UpDataCY
	VAR_INPUT
		Handle 	: UDINT;
	END_VAR
  VAR
  	p_SDO_act             : ^SDOHeader;
    us_SDO_length         : USINT;
    i                     : UINT;
    p_ReceiveObj          : pVirtualBase;
    p_SDOviaPath          : ^SDOviaPath;
    sd_retval             : DINT;
    IsStandardResp        : BOOL;
		SDORequestBuffer      : SDORequReadConfig;
    DataLen               : USINT;
    us_UnsafeSchedulerRun : USINT;
    p_PDOInBufferAct      : ^PDOInputBuffer;
    EverythingSynchron    : BOOL;
		MyPara 	              : CmdStruct;
		MyResult	            : results;
    UnsafeWrPackageNo     : USINT;
    aUnsafeWrPackages     : UnsafeWritePackages;
    UnsafeRdPackageNo     : USINT;
    aUnsafeRdPackages     : UnsafeReadPackages;
    TmpVal                : DINT;
    AddUnsafePackage      : BOOL;
    GotNewUnsafeValue     : BOOL;
    pHelpUnsafe           : ^UnsafeIORoutingElement;
    BDINTWriteVars        : USINT;
  END_VAR

//============================ Profiler start======================================================
#ifdef  DM_Profiler
  StartTimeMeasurement(usMode := DMTIME_CY);
#endif
//============================ Profiler end========================================================

  // do logging if necessary
  if bd_LogOnceMarker <> bd_AlreadyLoggedMarker then
    if bd_LogOnceMarker.MoveSourceInvalid > bd_AlreadyLoggedMarker.MoveSourceInvalid then
      bd_AlreadyLoggedMarker.MoveSourceInvalid := TRUE;
      LogError("@ZZZZ (SafetyCDIAS_Base::WritePDO2Module) [SL] Can't change Move-Command, because the new source address is invalid");
    end_if;

    if bd_LogOnceMarker.TdoLen0 > bd_AlreadyLoggedMarker.TdoLen0 then
      bd_AlreadyLoggedMarker.TdoLen0 := TRUE;
      LogError("@ZZZZ (SafetyCDIAS_Base::UpDateRT) [SL] Found TDOFrame with Length = 0");
    end_if;

    if bd_LogOnceMarker.TdoLenInvalid > bd_AlreadyLoggedMarker.TdoLenInvalid then
      bd_AlreadyLoggedMarker.TdoLenInvalid := TRUE;
      LogError("@ZZZZ (SafetyCDIAS_Base::UpDateRT) [SL] Found TDOFrame with invalid Length value inside (must be 20)");
    end_if;
  end_if;

  // do sdo communication only, if module has been found and initialized correctly and if there are some LEDs on (else a FW-Update is running)
  if ( State.uiIO_Flags = 0 ) & (VoltageOK | RunState | ServiceMode | Error) &
     (( ClassState = _SafetyClassOK ) | ( ClassState = _WaitForSynchronicity ) | ( ClassState = _ReinitConfig ) | ( ClassState = _ModFromCfgNotFound ) | ( ClassState = _UnknownCfgError ) | ( ClassState = _UnsafeVarNotFound )) then

    // wait until the safetymanager has initialized connection
    if b_ManagerReadyForSDO = FALSE then
      return;
    end_if;

    //Update of service messages doesn't take place in realtime

    // if we have to quit the communication errors and there is no other request open at this time
    if (QuitComError = 1) & (LastRequest = _NoOpenRequest) then
      if UnsafeScheduler <> UnsafeSchedulerSetBusReady then
        us_SetBusReadyState := WaitPDOsSyncron;
        UnsafeScheduler     := UnsafeSchedulerSetBusReady;
      end_if;

      QuitComError := 0;
    end_if;

    //read SDO from module and send it to the target module
    //check, if SDO is available and valid
    if ( p_Handle_SDO_Read^.us_Status = SAFETY_SDO_DATA_VALID ) then

      //calculate length of SDO
      us_SDO_length := sizeof(SDOHeader.StdHeader.CRC) + p_Handle_SDO_Read^.SDOStructure.SDOHeader.StdHeader.Len;

      //copy SDO without first byte (=status byte)
      To_StdLib.MemCpy(dest := p_SDOOutputBuffer, source := #p_Handle_SDO_Read^.SDOStructure, size := us_SDO_length );

#ifdef SAFETY_PROTOCOL_ANALYZER_ACTIVATED
  RecordFrame(p_SDOOutputBuffer$^DINT, 0);
#endif

      //mark data as received
      p_Handle_SDO_Read^.us_Status := SAFETY_SDO_NO_DATA;

      //find target object for routing
      p_ReceiveObj    := NIL;

      IsStandardResp  := FALSE;
      //check, if receiver is addressed by safety number or hardware path
      if ( (p_SDOOutputBuffer^.SDOHeader.StdHeader.Typ AND SSDO_MASK_TYPE) = FRM_TYPECODE_SSDO_MOD ) then

        //search this-pointer of receiver with safety number
        p_ReceiveObj := ( GetRoutingPointerByNumber(ud_SafeNumber := p_SDOOutputBuffer^.SDOHeader.DstAdr))$pVirtualBase;

      elsif ( (p_SDOOutputBuffer^.SDOHeader.StdHeader.Typ AND SSDO_MASK_TYPE) = FRM_TYPECODE_SSDO_MOD_TP ) then

        //search this-pointer of receiver with hardware path
        p_SDOviaPath := p_SDOOutputBuffer$^SDOviaPath;
        p_ReceiveObj := ( GetRoutingPointerByPath(p_ActObjectPath := #p_SDOviaPath^.TopologyPath[0], p_SDOviaPath^.StdHeader.Len - 8))$pVirtualBase;

      elsif ( (p_SDOOutputBuffer^.SDOHeader.StdHeader.Typ AND SSDO_MASK_TYPE) = FRM_TYPECODE_STD ) then
        IsStandardResp    := TRUE;
        StandardResponse  := (p_SDOOutputBuffer$^StandardFrameType)^;
        if StandardResponse.SDOHeader.SeqNr = (StandardSeqNr OR 16#80) then

          case LastRequest of
            _NoOpenRequest: // error, no open request, but we got a response
              LogError("@ZZZZ (SafetyCDIAS_Base::UpDataCY) Standard frame response received, without open request");

            _SetBusReady:
              IF StandardResponse.SDOHeader.Cmd = SDO_COMMAND_SET_BUS_READY THEN
                if us_SetBusReadyState <> SendSetBusReady then
                  LogError("@ZZZZ (SafetyCDIAS_Base::UpDataCY) Got Response of SetBusReady, but SSW is not in the right step");
                  return;
                end_if;
                us_SetBusReadyState := SetBusReadyFinished;
                b_ManualQuit    := FALSE;
                UnsafeScheduler := UnsafeSchedulerGetDiagVars; // Go on with the action-steps, done here so we don't lose a whole cycle
                LastRequest     := _NoOpenRequest;
                ud_AsyComRetryCounter := 0; // reset retry counter
                if ClassState = _WaitForSynchronicity then
                  ClassState    := _SafetyClassOK;
                end_if;
              else
                LogError("@ZZZZ (SafetyCDIAS_Base::UpDataCY) Invalid command: bus ready expected");
              END_IF;

            _ReadData:
              // if we did read command, then save the value to corresponding server
              if StandardResponse.SDOHeader.Cmd = SDO_COMMAND_READ then
                // if returncode is 0 read succeeded
                if StandardResponse.aData[0] = 0 then
                  // check if length is correct
                  if StandardResponse.aData[1] = StandardRequest.aData[4] then
                    // delete request
                    LastRequest := _NoOpenRequest;
                    ud_AsyComRetryCounter := 0; // reset retry counter

                    if (DiagVars.SavingLogSSW = GetLogFileBlocks) then
                      // save the last block in the memory for the file
                      _memcpy(ptr1:=DiagVars.pLogFileMem$pVoid + (DiagVars.LogHeader.LogMemSize - DiagVars.LogMemToGet),
                              ptr2:=#StandardResponse.aData[2],
                              cntr:=DiagVars.BytesToGet);

                      DiagVars.LogMemToGet -= DiagVars.BytesToGet;

                      if DiagVars.LogMemToGet = 0 then
                        DiagVars.SavingLogSSW := GetLogHeader2;
                      end_if;
                    else
                      LogError("@ZZZZ (SafetyCDIAS_Base::UpDataCY) SDO Receive: Invalid Read response (no diagnostic read active)");
                    end_if;
                  end_if;
                end_if;
              else
                LogError("@ZZZZ (SafetyCDIAS_Base::UpDataCY) SDO Receive: Invalid command, read expected");
              end_if;

            _ReadValues:
              // if we did read command, then save the value to corresponding server
              if StandardResponse.SDOHeader.Cmd = SDO_COMMAND_READ_VALUES then
                // if returncode is 0 read succeeded
                if StandardResponse.aData[0] = 0 then
                  // check if length is correct
                  if StandardResponse.aData[1] = StandardRequest.aData[0] then
                    // delete request
                    LastRequest := _NoOpenRequest;
                    ud_AsyComRetryCounter := 0; // reset retry counter

                    // if we got some outputs in the routing table and a valid pointer, write values to servers
                    if ui_CntUnsafeOutputs & pUnsafeOutElement then

                      // depending on length we do different number of server write-methods to set the data we just read
//                      pUnsafeOutElement := p_UnsafeOutputsTable + (UnsafeReadTransNr * MaxVarsPerReadPackage * sizeof(UnsafeIORoutingElement));  // the pointer is already on this element
                      for i := 0 to (StandardResponse.aData[1] - 1) do
                        // save the new value temporarily
                        TmpVal := StandardResponse.aData[2 + (i * sizeof(DINT))]$DINT;
                        if pUnsafeOutElement^.ud_Thisp then
                          if pUnsafeOutElement^.UnsafeType = BDINTOutput then
                            pUnsafeOutElement^.sd_OldValue := RD(pUnsafeOutElement^.ud_Thisp$^void)$DINT;
                            TmpVal := ((pUnsafeOutElement^.sd_OldValue$UDINT AND (NOT pUnsafeOutElement^.BitMask)) OR
                                      (TmpVal$UDINT AND pUnsafeOutElement^.BitMask))$DINT;

                            // now we have to write the value to the server
                            WR(pUnsafeOutElement^.ud_Thisp$^void, TmpVal);
                          else
                            WR(pUnsafeOutElement^.ud_Thisp$^void, TmpVal);
                          end_if;
                        elsif (pUnsafeOutElement^.UnsafeType = ExternalOutput) | (pUnsafeOutElement^.UnsafeType = ExternalBDINTOutput) then
                          pUnsafeOutElement^.sd_NewValue4External := TmpVal;

                          // mark the value as valid
                          pUnsafeOutElement^.b_IsValid := TRUE;
                        end_if;
                        pUnsafeOutElement += sizeof(UnsafeIORoutingElement);
                      end_for;
                    end_if;

                    UnsafeReadTransNr += 1;
                  end_if;
                end_if;
              else
                LogError("@ZZZZ (SafetyCDIAS_Base::UpDataCY) SDO Receive: Invalid command, read values expected");
              end_if;

            _WriteValues:
              if IsOptimizedCPU() then
                // if we did a write command, just check
                if StandardResponse.SDOHeader.Cmd = SDO_COMMAND_WRITE_VALUES then
                  // delete request
                  LastRequest := _NoOpenRequest;
                  ud_AsyComRetryCounter := 0; // reset retry counter

                  // if there is no more element to send or check for changes => proceed to the next step
                  if pUnsafeInElement = NIL then
                    UnsafeScheduler := UnsafeSchedulerReadData; //We need to set scheduler to next step....
                  end_if;
                else
                  LogError("@ZZZZ (SafetyCDIAS_Base::UpDataCY) SDO Receive: Invalid command, write expected");
                end_if;
              else
                // on CSCP011 the SDO_COMMAND_WRITE_VALUES didn't exist

                // if we did a write command, just check
                if StandardResponse.SDOHeader.Cmd = SDO_COMMAND_WRITE then
                  // delete request
                  LastRequest           := _NoOpenRequest;
                  ud_AsyComRetryCounter := 0; // reset retry counter

                  if UnsafeWriteTransNr < (WriteFramesNeeded - 1) then
                    UnsafeWriteTransNr  += 1;
                  else
                    UnsafeWriteTransNr  := 0;
                    UnsafeWritingActive := FALSE;
                    UnsafeScheduler     := UnsafeSchedulerReadData; //We need to set scheduler to next step....
                  end_if;
                else
                  LogError("@ZZZZ (SafetyCDIAS_Base::UpDataCY) SDO Receive: Invalid command, write expected");
                end_if;
              end_if;

            _GetCRC:
              // check if it's a response to a read command
              if StandardResponse.SDOHeader.Cmd = SDO_COMMAND_READ then
                // if returncode is 0 read succeeded
                if StandardResponse.aData[0] = 0 then
                  // check if length is correct
                  if StandardResponse.aData[1] = 4 then

                    // delete request
                    LastRequest := _NoOpenRequest;
                    ud_AsyComRetryCounter := 0; // reset retry counter

                    if ud_ConfigCRC <> StandardResponse.aData[2]$UDINT then
                      // CRC has changed => save the new crc
                      ud_ConfigCRC          := StandardResponse.aData[2]$UDINT;
                      //Show CRC on Server
                      DesignerPrjConfigCRC  := ud_ConfigCRC;

                      // show that we read the config of the class again
                      ClassState            := _ReinitConfig;

                      if pSafetyManagerThis then
                        MyPara.uiCmd    := CMD_SM_NEW_SAFETY_PROJECT;
                        MyPara.aPara[0] := 4;
                        MyPara.aPara[4] := (#SafetyNumber)$DINT;
                        pSafetyManagerThis^.NewInst(#MyPara, #MyResult);
                      end_if;

                      // remove the cpu from all classes, which use it
                      ResetConfig();

                      // we have to return here because:
                      // the command CMD_SM_NEW_SAFETY_PROJECT will trigger a disconnect of this class which will set the unsafe scheduler to setbusready,
                      // which would skip the synchron check in the actual cyclic run because everything of the old configuration is synchron now
                      return;
                    end_if;
                  end_if;
                end_if;
              end_if;

            _DiagState:
              if StandardResponse.SDOHeader.Cmd = SDO_COMMAND_GET_STATE then
                _memcpy(ptr1 := #DiagVars.UserGetStateResp,
                        ptr2 := #StandardResponse.aData + SIZEOF(USINT),
                        cntr := sizeof(GetStateResponseType) );
                DiagVars.UserDiagStateReady := TRUE;
                DiagVars.UserWantsDiagState := FALSE;
                LastRequest                 := _NoOpenRequest;
                ud_AsyComRetryCounter       := 0; // reset retry counter
              end_if;
            _DiagInfo:
              if StandardResponse.SDOHeader.Cmd = SDO_COMMAND_GET_DIAG_INFO then
                _memcpy(ptr1 := #DiagVars.UserGetDiagInfoResp,
                        ptr2 := #StandardResponse.aData + SIZEOF(USINT),
                        cntr := sizeof(SafetyDiagInfo) );
                DiagVars.UserDiagInfoReady  := TRUE;
                DiagVars.UserWantsDiagInfo  := FALSE;
                LastRequest                 := _NoOpenRequest;
                ud_AsyComRetryCounter       := 0; // reset retry counter
              end_if;

            _ErrorChannelInfo:
            //if we did read command, then save the value to corresponding server
              if StandardResponse.SDOHeader.Cmd = SDO_COMMAND_READ then
                // if returncode is 0 read succeeded
                if StandardResponse.aData[0] = 0 then
                  // check if length is correct
                  if StandardResponse.aData[1] <> 0  then
                    _memcpy(ptr1 := #aErrorMem[actoffset],
                            ptr2 := #StandardResponse.aData[2],
                            cntr := StandardResponse.aData[1]);
                    if remainingPacketlength = 0 then
                      remainingPacketlength := StandardResponse.aData[2] - StandardResponse.aData[1];
                      actoffset := StandardResponse.aData[1];
                    else
                      remainingPacketlength -= StandardResponse.aData[1];
                      actoffset += StandardResponse.aData[1];
                    end_if;

                    // delete request
                    LastRequest := _NoOpenRequest;
                    if remainingPacketlength <= 0  then
                      //Finish reset variables
                      DiagVars.UserErrorInfoReady := TRUE;
                      DiagVars.UserWantsErrorInfo := FALSE;
                      ud_AsyComRetryCounter := 0; // reset retry counter
                      remainingPacketlength := 0; //reset remainingPacketlength
                      actoffset := 0; //reset offset
                    end_if;
                  end_if;
                end_if;
              end_if;
          else
            LogError("@ZZZZ (SafetyCDIAS_Base::UpDataCY) SDO Receive: Invalid standard frame response");
          end_case;

          // if request is deleted, increase sequence number to set next request
          if LastRequest = _NoOpenRequest then
            if StandardSeqNr < 16#7F then
              StandardSeqNr += 1;
            else
              StandardSeqNr := 0;
            end_if;
          end_if;
        else
          LogError("@ZZZZ (SafetyCDIAS_Base::UpDataCY) SDO Receive: Invalid sequence number in Standard SDO response");
          LogValue("expected: {0} / received: {1}", Value:=(StandardSeqNr OR 16#80), Value2:=StandardResponse.SDOHeader.SeqNr);
        end_if;
      else
        LogError("@ZZZZ (SafetyCDIAS_Base::UpDataCY) SDO Receive: Invalid frametype in Standard SDO response");
      end_if;

      // dont let the CDIAS-modules start before the master-slave configuation has finished (don´t forward the GetState to itself)
      if (p_ReceiveObj = this) & (b_ManagerInitialisationFinished = FALSE) then
        case ud_MyModuleID of
          CSCP01x_ID,
          CSDI16x_ID,
          CSTO08x_ID:
            // set some flags to ignore the SDO
            p_ReceiveObj    := NIL;
            IsStandardResp  := TRUE;
        end_case;
      end_if;

      //if there is no object, the message will be lost
      if ( p_ReceiveObj ) then

        //send SDO to receiver object
        MyPara.uiCmd    := CMD_SM_ADD_SDO_TO_BUFFER;
        MyPara.aPara[0] := p_SDOOutputBuffer$DINT;
        MyPara.aPara[1] := us_SDO_length;
        sd_retval$iprStates := p_ReceiveObj^.NewInst(#MyPara, #MyResult);

//        sd_retval := p_ReceiveObj^.AddSDOToBuffer(p_us_Message := p_SDOOutputBuffer$^USINT, us_length := us_SDO_length);

        if sd_retval then
          // generate error message with returncode (add to logfile and debugger trace)
          LogValue("@ZZZZ (SafetyCDIAS_Base::UpDataCY) AddSDOToBuffer failed: Returncode: -0x{0}", Value:=(0-sd_retval)$UDINT);
        end_if;

      elsif IsStandardResp = FALSE then

        if pSafetyManagerThis & us_SDO_length then
#ifdef DO_DEBUG
          DOCheck(pFrame:=(p_SDOOutputBuffer)$^SDOStdHeader, pCheckStruct:=#SDORead);
#endif

          MyPara.uiCmd    := CMD_SM_SDO_TO_MANAGER;
          MyPara.aPara[0] := to_dint(us_SDO_length);
          MyPara.aPara[1] := p_SDOOutputBuffer$DINT;
          pSafetyManagerThis^.NewInst(#MyPara, #MyResult);
        else
          //log not routable SDOs
          LogValue("@ZZZZ (SafetyCDIAS_Base::UpDataCY) Safety module {0}: SDO not routed to receiver {1}", SafetyNumber$UDINT, p_SDOOutputBuffer^.SDOHeader.DstAdr$UDINT);
        end_if;
      end_if;

    elsif (LastRequest <> _NoOpenRequest) & (ud_TransfertimePerPackage > 0) then
      // count up for timeout
      ud_UnsafeTimeoutCounter += 1;

      if ( ud_UnsafeTimeoutCounter ) > ( 50 * ud_TransfertimePerPackage ) then
        CASE UnsafeScheduler OF

          UnsafeSchedulerSetBusReady:
            LogError("@ZZZZ (SafetyCDIAS_Base::UpdateCy) Timeout on setting bus ready");

          UnsafeSchedulerGetDiagVars:
            IF LastRequest = _ReadData THEN
              LogError("@ZZZZ (SafetyCDIAS_Base::UpdateCy) Timeout requesting DiagVars");
            END_IF;
            UnsafeScheduler       := UnsafeSchedulerGetCRC;
            DiagVars.SavingLogSSW := GetLogFileBlocks;

          UnsafeSchedulerGetCRC:
            LogError("@ZZZZ (SafetyCDIAS_Base::UpdateCy) Timeout requesting CRC");
            UnsafeScheduler       := UnsafeSchedulerWriteData;

          UnsafeSchedulerWriteData:
            LogError("@ZZZZ (SafetyCDIAS_Base::UpdateCy) Timeout writing Data 'Unsafe Input'");
            UnsafeScheduler       := UnsafeSchedulerReadData;
            UnsafeWriteTransNr    := 0;

          UnsafeSchedulerReadData:
            LogError("@ZZZZ (SafetyCDIAS_Base::UpdateCy) Timeout reading Data 'Unsafe Output'");
            UnsafeScheduler       := UnsafeSchedulerDiagState;
            UnsafeReadTransNr     := 0;

          UnsafeSchedulerDiagState:
            LogError("@ZZZZ (SafetyCDIAS_Base::UpdateCy) Timeout on reading DiagState");
            UnsafeScheduler       := UnsafeSchedulerDiagInfo;

          UnsafeSchedulerDiagInfo:
            LogError("@ZZZZ (SafetyCDIAS_Base::UpdateCy) Timeout on reading DiagInfo");
            UnsafeScheduler       := UnsafeSchedulerChannelError;

          UnsafeSchedulerChannelError:
            LogError("@ZZZZ (SafetyCDIAS_Base::UpdateCy) Timeout on reading ChannelError");
            UnsafeScheduler       := UnsafeSchedulerGetDiagVars;

        END_CASE;

        // we only increase the retry counter if the module is running
        if RunState then
          ud_AsyComRetryCounter += 1;
        end_if;

        if ud_AsyComRetryCounter >= SDO_MAX_TRIES then
          ClassState := _AsyncComError;
          LogError("@ZZZZ (SafetyCDIAS_Base::UpdateCy) Too many consecutive asynchronous commands failed! Please contact Sigmatek Support!");
        else
          LastRequest := _NoOpenRequest;
          // if request is deleted, increase sequence number to set next request
          if StandardSeqNr < 16#7F then
            StandardSeqNr += 1;
          else
            StandardSeqNr := 0;
          end_if;
        end_if;
      end_if;

    end_if;

    //write to hardware from other module received SDO
    if ( ui_cnt_SDOInputBuffer > 0 ) & p_SDOInputBuffer then

      //set pointer to first SDO in the SDO list
      p_SDO_act     := p_SDOInputBuffer$^SDOHeader;

      //calculate length of SDO (CRC + data length)
      us_SDO_length := sizeof (SDOHeader.StdHeader.CRC) + p_SDO_act^.StdHeader.Len;

      //check, if buffer is empty
      if ( p_Handle_SDO_Write^.us_Status = SAFETY_SDO_NO_DATA ) then

#ifdef SAFETY_PROTOCOL_ANALYZER_ACTIVATED
  RecordFrame(p_SDO_act$^DINT, 1);
#endif

        //copy SDO into write-buffer
        To_StdLib.MemCpy(dest := #p_Handle_SDO_Write^.SDOStructure, source := p_SDO_act, size := us_SDO_length);

        //mark SDO data as valid
        p_Handle_SDO_Write^.us_Status := SAFETY_SDO_DATA_VALID;

        //decrement amount of SDOs
        ui_cnt_SDOInputBuffer -= 1;

        //if there is at least 1 SDO left, copy the remaining memory over the actual SDO
        if ( ui_cnt_SDOInputBuffer > 0 ) then

          //remove first entry in the SDO list
          _memmove(p_SDOInputBuffer, (p_SDOInputBuffer + SDO_MAX_LENGTH), (ui_cnt_SDOInputBuffer * SDO_MAX_LENGTH));
        end_if;
      end_if;
    end_if;

    // Start of scheduler; we need to share the time between reading, writing and diagnosis
    us_UnsafeSchedulerRun := 0;

    if (b_ManagerInitialisationFinished = TRUE) & ( ClassState <> _ReinitConfig ) & ( p_Handle_SDO_Write^.us_Status = SAFETY_SDO_NO_DATA ) then

      // Check actions until we find somthing we need to do
      // all 6 action-steps must be walked through during one cycle to make sure new data is fetched as fast as possible
      // SetBusReady is an exception: this step is only performed once on bootup!
      while (us_UnsafeSchedulerRun < 6) & (LastRequest = _NoOpenRequest) do
        us_UnsafeSchedulerRun   += 1;
        ud_UnsafeTimeoutCounter := 0; //No active request: we can reset the timeout-counter
        case UnsafeScheduler of

       (* ***************************************** *)
          UnsafeSchedulerSetBusReady:
       (* ***************************************** *)
          case us_SetBusReadyState of

          //-------------------------------------------------------------------------------------------------------------
            WaitPDOsSyncron:

              EverythingSynchron := TRUE;

              // it's possible that all PDOs are coming from a different domain, then we have no inputbuffer
              if ui_cnt_PDOInputBuffer then
                p_PDOInBufferAct := #aPDOInputBuffer[0];
                for i := 0 to (ui_cnt_PDOInputBuffer-1) do
                  if p_PDOInBufferAct^.b_TimeSynchron = FALSE then
                    // we're still not synchron with this module. if it's optional it is probably not connected
                    if p_PDOInBufferAct^.b_IsOptional then
                      if (ops.tAbsolute - ud_OptionalTimeoutStart) <= OPTIONAL_MODULE_SYNC_TIMEOUT then
                        // if timeout not exceeded => not sychron (otherwise the variable will stay on it's old value)
                        EverythingSynchron  := FALSE;
                        exit;
                      else
                        TRACE("Synchronisation timeout for optional module exceeded => assume it's synchon");
                      end_if;
                    else
                      EverythingSynchron    := FALSE;
                      exit;
                    end_if;
                  end_if;

                  p_PDOInBufferAct +=  sizeof(PDOInputBuffer);
                end_for;

                if EverythingSynchron & (ModuleSyncNo > 0) then
                  ModuleSyncNo -= 1;

#ifdef SAFETY_DEBUG_LOGGING_ACTIVATED
//                  case ud_MyModuleID of
//                    CSCP01x_ID:
//                      TRACE("ModuleSyncNo wurde dekrementiert von: CSCP");
//
//                    CSDI16x_ID:
//                      TRACE("ModuleSyncNo wurde dekrementiert von: CSDI");
//
//                    CSTO08x_ID:
//                      TRACE("ModuleSyncNo wurde dekrementiert von: CSTO");
//                  end_case;
#endif
                end_if;
#ifdef SAFETY_DEBUG_LOGGING_ACTIVATED
//              elsif EverythingSynchron then
//                  case ud_MyModuleID of
//                    CSCP01x_ID:
//                      TRACE("ModuleSyncNo wurde nicht verändert von: CSCP");
//
//                    CSDI16x_ID:
//                      TRACE("ModuleSyncNo wurde nicht verändert von: CSDI");
//
//                    CSTO08x_ID:
//                      TRACE("ModuleSyncNo wurde nicht verändert von: CSTO");
//                  end_case;
#endif
              end_if;

              if EverythingSynchron then
                us_SetBusReadyState := WaitAllModulesSyncron;
              end_if;

          //-------------------------------------------------------------------------------------------------------------
            WaitAllModulesSyncron:
              // wait for other modules to be synchron with each other
              if (ModuleSyncNo = 0) & b_ManagerInitialisationFinished then
                us_SetBusReadyState := SendSetBusReady;
              end_if;

          //-------------------------------------------------------------------------------------------------------------
            SendSetBusReady:
              // send the bus-ready command
              SDORequestBuffer.StdHeader.CRC  := 0;                                                   // CRC is always 0 in Std communication
              SDORequestBuffer.StdHeader.Cmd  := SDO_COMMAND_SET_BUS_READY;                           // set bus ready command
              SDORequestBuffer.StdHeader.Typ  := FRM_TYPECODE_STD;                                    // standard frame type
              SDORequestBuffer.StdHeader.SeqNr:= StandardSeqNr OR 16#80;                              // sequence number
              SDORequestBuffer.StdHeader.Len  := 4;                                                   // header

              LastRequest := _SetBusReady;

#ifdef SAFETY_PROTOCOL_ANALYZER_ACTIVATED
  RecordFrame((#SDORequestBuffer)$^DINT, 1);
#endif

              //copy SDO into write-buffer
              To_StdLib.MemCpy(dest := #p_Handle_SDO_Write^.SDOStructure, source := #SDORequestBuffer, size := (sizeof(SDOHeader.StdHeader.CRC) + SDORequestBuffer.StdHeader.Len));

              //mark SDO data as valid
              p_Handle_SDO_Write^.us_Status := SAFETY_SDO_DATA_VALID;

              if ( pISafety^.udVersion >= 16#1001 ) then
                SAFETY_iPushSafetyTask();
              end_if;

          //-------------------------------------------------------------------------------------------------------------
            SetBusReadyFinished:
              // all ok, nothing to do here

          end_case;
          us_UnsafeSchedulerRun := 16#FF; //make sure we don't repeat the while-loop until we have sent the bus-ready command

       (* ***************************************** *)
          UnsafeSchedulerGetDiagVars:
       (* ***************************************** *)

          //check, if buffer is empty and we got some unsafe data to get/set and crc check is finished
          if (DiagVars.SavingLogSSW = GetLogFileBlocks) then

            // check if more than blocksize to get
            if DiagVars.LogMemToGet > LOG_DATA_BLOCK_SIZE then
              // get a complete block
              DiagVars.BytesToGet := LOG_DATA_BLOCK_SIZE;
            else
              // get only the last bytes
              DiagVars.BytesToGet := DiagVars.LogMemToGet$USINT;
            end_if;

            StandardRequest.SDOHeader.Cmd   := SDO_COMMAND_READ;                            // read command
            StandardRequest.SDOHeader.Typ   := FRM_TYPECODE_STD;                            // standard frame type
            StandardRequest.SDOHeader.SeqNr := StandardSeqNr OR 16#80;                      // sequence number is in special area
            StandardRequest.SDOHeader.Len   := 4 + 4 + 1;                                   // header + destination address + length of data
            StandardRequest.aData[0]$UDINT  := DiagVars.ReadBaseAdr + (DiagVars.LogHeader.LogMemSize - DiagVars.LogMemToGet);// destination address
            StandardRequest.aData[4]        := DiagVars.BytesToGet$USINT;                   // length of data

            LastRequest := _ReadData;

#ifdef SAFETY_PROTOCOL_ANALYZER_ACTIVATED
  RecordFrame((#StandardRequest)$^DINT, 1);
#endif

            //copy SDO into write-buffer
            To_StdLib.MemCpy(dest := #p_Handle_SDO_Write^.SDOStructure, source := #StandardRequest, size := (sizeof(SDOHeader.StdHeader.CRC) + StandardRequest.SDOHeader.Len));

            //mark SDO data as valid
            p_Handle_SDO_Write^.us_Status := SAFETY_SDO_DATA_VALID;

            if ( pISafety^.udVersion >= 16#1001 ) then
              SAFETY_iPushSafetyTask();
            end_if;
          else
            UnsafeScheduler := UnsafeSchedulerGetCRC;
          end_if;

       (* ***************************************** *)
          UnsafeSchedulerGetCRC:
       (* ***************************************** *)

          // every 5 secs check for a new safety project inside the cpu
          if b_CheckCRC & ((ops.tAbsolute - ud_LastCrcCheck) > CRC_CHECK_TIME ) then

            SDORequestBuffer.StdHeader.CRC  := 0;                                                   // CRC is always 0 in Std communication
            SDORequestBuffer.StdHeader.Cmd  := SDO_COMMAND_READ;                                    // read command
            SDORequestBuffer.StdHeader.Typ  := FRM_TYPECODE_STD;                                    // standard frame type
            SDORequestBuffer.StdHeader.SeqNr:= StandardSeqNr OR 16#80;                              // sequence number
            SDORequestBuffer.StdHeader.Len  := 4 + 4 + 1;                                           // header + destination address + length of data
            SDORequestBuffer.ud_Address     := SDO_ADDRESS_CONFIG_DATA + SDO_OFFSET_CONFIG_CRC_ALL; // address of crc
            SDORequestBuffer.us_Length      := 4;                                                   // length of crc

            LastRequest := _GetCRC;

#ifdef SAFETY_PROTOCOL_ANALYZER_ACTIVATED
  RecordFrame((#SDORequestBuffer)$^DINT, 1);
#endif

            //copy SDO into write-buffer
            To_StdLib.MemCpy(dest := #p_Handle_SDO_Write^.SDOStructure, source := #SDORequestBuffer, size := (sizeof(SDOHeader.StdHeader.CRC) + SDORequestBuffer.StdHeader.Len));

            //mark SDO data as valid
            p_Handle_SDO_Write^.us_Status := SAFETY_SDO_DATA_VALID;

            if ( pISafety^.udVersion >= 16#1001 ) then
              SAFETY_iPushSafetyTask();
            end_if;

            ud_LastCrcCheck := ops.tAbsolute;
          else
            if RunState then
              // in operational also get unsave-variables
              UnsafeScheduler := UnsafeSchedulerWriteData;
            else
              // not operational, we must skip the unsave vars
              UnsafeScheduler := UnsafeSchedulerDiagState;
              us_UnsafeSchedulerRun += 2;
            end_if;
          end_if;

       (* ***************************************** *)
          UnsafeSchedulerWriteData:
       (* ***************************************** *)

          if IsOptimizedCPU() then
            if ui_CntUnsafeInputs then
              // if we have finished checking through all variables the last time => check from beginning (otherwise the pointer is on the element where we have to continue)
              if pUnsafeInElement = NIL then
                pUnsafeInElement := p_UnsafeInputsTable;
              end_if;

              // we check if we have to write any of the unsafe input variables (only until our message is full)
              UnsafeWrPackageNo := 0;
              BDINTWriteVars    := 0; // limit number of bdint write variables to 3 to ensure constant load of firmware
              while pUnsafeInElement & (UnsafeWrPackageNo < MAX_UNSAFE_WRITE_PACKAGES) & (BDINTWriteVars < MAX_UNSAFE_BDINTS_PER_WRITE) do

                // we have to check if we add this one
                GotNewUnsafeValue := FALSE;

                // if the type is normal we can read the actual value from the server
                if pUnsafeInElement^.UnsafeType = NormalUnsafe then
                  // check if pointer to server is valid
                  if pUnsafeInElement^.ud_Thisp then
                    // get the actual value from the server
                    TmpVal := RD((pUnsafeInElement^.ud_Thisp)$^void);

                    // we remember to update this if it's necessary
                    GotNewUnsafeValue := TRUE;
                  else
                    if bd_LogOnceMarker.NoThisForUnsafeIn = FALSE then
                      bd_LogOnceMarker.NoThisForUnsafeIn        := TRUE;
                      bd_AlreadyLoggedMarker.NoThisForUnsafeIn  := TRUE;
                      LogError("@ZZZZ (SafetyCDIAS_Base::UpdateCy) [SL] No thispointer available for Server of local unsafe input variable");
                    end_if;
                  end_if;
                elsif pUnsafeInElement^.UnsafeType = ExternalInput then
                  // check if we already have a valid value there
                  if pUnsafeInElement^.b_IsValid then
                    // get the actual value from the element
                    TmpVal := pUnsafeInElement^.sd_NewValue4External;

                    // we remember to update this if it's necessary
                    GotNewUnsafeValue := TRUE;
                  end_if;
                else
                  if bd_LogOnceMarker.WrongUnsafeVarType = FALSE then
                    bd_LogOnceMarker.WrongUnsafeVarType       := TRUE;
                    bd_AlreadyLoggedMarker.WrongUnsafeVarType := TRUE;
                    LogError("@ZZZZ (SafetyCDIAS_Base::UpdateCy) [SL] Wrong unsafe variable type in unsafe input list");
                  end_if;
                end_if;

                // if we have a new valid unsafe value => check if we have to send it
                if GotNewUnsafeValue then
                  // if it hasn't been sent yet
                  if (pUnsafeInElement^.b_AlreadyTransmitted = FALSE) then
                    // remember that we sent this already
                    pUnsafeInElement^.b_AlreadyTransmitted := TRUE;

                    // add this one
                    AddUnsafePackage := TRUE;
                  elsif TmpVal <> pUnsafeInElement^.sd_OldValue then
                    // if there were any changes on this value

                    // add this one
                    AddUnsafePackage := TRUE;
                  else
                    // don't add this one
                    AddUnsafePackage := FALSE;
                  end_if;

                  // if it is ready to be added => add it to send buffer
                  if AddUnsafePackage then
                    // add a package to send
                    aUnsafeWrPackages[UnsafeWrPackageNo].ud_Address := pUnsafeInElement^.ud_Address;
                    aUnsafeWrPackages[UnsafeWrPackageNo].Value      := TmpVal;
                    UnsafeWrPackageNo += 1;

                    // if it has a bitmask it's an unsafe bdint input variable
                    if pUnsafeInElement^.BitMask then
                      BDINTWriteVars += 1;
                    end_if;

                    // remember the actual as old value
                    pUnsafeInElement^.sd_OldValue := TmpVal;
                  end_if;
                end_if;

                pUnsafeInElement := pUnsafeInElement^.pNext;
              end_while;

              if UnsafeWrPackageNo then
                DataLen := UnsafeWrPackageNo * sizeof(UnsafeWritePackage);

                StandardRequest.SDOHeader.Cmd                 := SDO_COMMAND_WRITE_VALUES;       // write values command
                StandardRequest.SDOHeader.Typ                 := FRM_TYPECODE_STD;               // standard frame type
                StandardRequest.SDOHeader.SeqNr               := StandardSeqNr OR 16#80;         // sequence number is in special area
                StandardRequest.SDOHeader.Len                 := 4 + 4 + 1 + DataLen;            // header + destination address + length of data + data
                StandardRequest.aData[0]                      := UnsafeWrPackageNo;              // number of packages
                StandardRequest.aData[1]$UnsafeWritePackages  := aUnsafeWrPackages;              // packages

                LastRequest := _WriteValues;

#ifdef SAFETY_PROTOCOL_ANALYZER_ACTIVATED
  RecordFrame((#StandardRequest)$^DINT, 1);
#endif

                //copy SDO into write-buffer
                To_StdLib.MemCpy(dest := #p_Handle_SDO_Write^.SDOStructure, source := #StandardRequest, size := (sizeof(SDOHeader.StdHeader.CRC) + StandardRequest.SDOHeader.Len));

                //mark SDO data as valid
                p_Handle_SDO_Write^.us_Status := SAFETY_SDO_DATA_VALID;

                if ( pISafety^.udVersion >= 16#1001 ) then
                  SAFETY_iPushSafetyTask();
                end_if;
              else
                UnsafeScheduler := UnsafeSchedulerReadData;
              end_if;
            else
              UnsafeScheduler   := UnsafeSchedulerReadData;
            end_if;
          else
            // on CSCP011 the SDO_COMMAND_WRITE_VALUES didn't exist
            if ui_CntUnsafeInputs & WriteFramesNeeded then
              // if writing is not active, check if it's necessary to activate it
              if (UnsafeWritingActive = FALSE) then
                pUnsafeInElement := p_UnsafeInputsTable;

                for i := 0 to (ui_CntUnsafeInputs - 1) do
                  if pUnsafeInElement^.ud_Thisp then
                    sd_retval := RD((pUnsafeInElement^.ud_Thisp)$^void);        // data
                    if pUnsafeInElement^.sd_OldValue <> sd_retval then
                      UnsafeWritingActive := TRUE;
                      pUnsafeInElement^.sd_OldValue := sd_retval;
                    end_if;
                  end_if;
                  pUnsafeInElement += sizeof(UnsafeIORoutingElement);
                end_for;
              end_if;

              // check if writing is already active
              if UnsafeWritingActive then
                // pointer to the right unsafe input
                pUnsafeInElement := p_UnsafeInputsTable + (UnsafeWriteTransNr * MaxVarsPerWritePackage * sizeof(UnsafeIORoutingElement));

                // get length of data we write
                if (UnsafeWriteTransNr < (WriteFramesNeeded-1)) | ((ui_CntUnsafeInputs MOD MaxVarsPerWritePackage) = 0) then
                  DataLen := MaxVarsPerWritePackage * sizeof(DINT);
                else
                  DataLen := (ui_CntUnsafeInputs MOD MaxVarsPerWritePackage)$USINT * sizeof(DINT);
                end_if;

                StandardRequest.SDOHeader.Cmd   := SDO_COMMAND_WRITE;                           // write command
                StandardRequest.SDOHeader.Typ   := FRM_TYPECODE_STD;                            // standard frame type
                StandardRequest.SDOHeader.SeqNr := StandardSeqNr OR 16#80;                      // sequence number is in special area
                StandardRequest.SDOHeader.Len   := 4 + 4 + 1 + DataLen;                         // header + destination address + length of data + data
                StandardRequest.aData[0]$UDINT  := pUnsafeInElement^.ud_Address;                // destination address
                StandardRequest.aData[4]        := DataLen;                                     // length of data

                // depending on length we do different number of server read-methods to get the data we write
                for i := 0 to (DataLen/sizeof(DINT)) - 1 do
                  if pUnsafeInElement^.ud_Thisp then
                    StandardRequest.aData[5 + (i * sizeof(DINT))]$DINT := pUnsafeInElement^.sd_OldValue;
                  else
                    // this server doesn't exist in lasal => always send 0
                    StandardRequest.aData[5 + (i * sizeof(DINT))]$DINT := 0;
                  end_if;

                  pUnsafeInElement += sizeof(UnsafeIORoutingElement);
                end_for;

                LastRequest := _WriteValues;

#ifdef SAFETY_PROTOCOL_ANALYZER_ACTIVATED
  RecordFrame((#StandardRequest)$^DINT, 1);
#endif

                //copy SDO into write-buffer
                To_StdLib.MemCpy(dest := #p_Handle_SDO_Write^.SDOStructure, source := #StandardRequest, size := (sizeof(SDOHeader.StdHeader.CRC) + StandardRequest.SDOHeader.Len));

                //mark SDO data as valid
                p_Handle_SDO_Write^.us_Status := SAFETY_SDO_DATA_VALID;

                if ( pISafety^.udVersion >= 16#1001 ) then
                  SAFETY_iPushSafetyTask();
                end_if;
              else
                UnsafeScheduler := UnsafeSchedulerReadData;
              end_if;
            else
              UnsafeScheduler   := UnsafeSchedulerReadData;
            end_if;
          end_if;

       (* ***************************************** *)
          UnsafeSchedulerReadData:
       (* ***************************************** *)
          if ui_CntUnsafeOutputs & ReadFramesNeeded then
            //check, if buffer is empty and we got some unsafe data to get/set and crc check is finished
            if (UnsafeReadTransNr < ReadFramesNeeded) //then
             & ( ((UnsafeReadTransNr = 0) & ( ops.tAbsolute - LastUnsafeUpdate > ud_ServerUpdateTime ) ) | (UnsafeReadTransNr <> 0) )then
              // here we request directly the unsafe IOs

              // sequence number is in special area
              StandardRequest.SDOHeader.SeqNr := StandardSeqNr OR 16#80;

              // we get an output
              pUnsafeOutElement := p_UnsafeOutputsTable + (UnsafeReadTransNr * MaxVarsPerReadPackage * sizeof(UnsafeIORoutingElement));

              // get length of data we read
              if (UnsafeReadTransNr < (ReadFramesNeeded - 1)) | ((ui_CntUnsafeOutputs MOD MaxVarsPerReadPackage) = 0) then
                UnsafeRdPackageNo := MaxVarsPerReadPackage;
              else
                UnsafeRdPackageNo := (ui_CntUnsafeOutputs MOD MaxVarsPerReadPackage)$USINT;
              end_if;

              DataLen := UnsafeRdPackageNo * sizeof(DINT);

              // create buffer with addresses of values to read
              pHelpUnsafe := pUnsafeOutElement;
              for i := 0 to (UnsafeRdPackageNo-1) do
                aUnsafeRdPackages[i] := pHelpUnsafe^.ud_Address;
                pHelpUnsafe += sizeof(UnsafeIORoutingElement);
              end_for;

              StandardRequest.SDOHeader.Cmd               := SDO_COMMAND_READ_VALUES;                     // read values command
              StandardRequest.SDOHeader.Typ               := FRM_TYPECODE_STD;                            // standard frame type
              StandardRequest.SDOHeader.SeqNr             := StandardSeqNr OR 16#80;                      // sequence number is in special area
              StandardRequest.SDOHeader.Len               := 4 + 1 + DataLen;                             // header + size + length of data
              StandardRequest.aData[0]                    := UnsafeRdPackageNo;                           // number of values to get
              StandardRequest.aData[1]$UnsafeReadPackages := aUnsafeRdPackages;                           // read addresses

              LastRequest := _ReadValues;

#ifdef SAFETY_PROTOCOL_ANALYZER_ACTIVATED
  RecordFrame((#StandardRequest)$^DINT, 1);
#endif

              //copy SDO into write-buffer
              To_StdLib.MemCpy(dest := #p_Handle_SDO_Write^.SDOStructure, source := #StandardRequest, size := (sizeof(SDOHeader.StdHeader.CRC) + StandardRequest.SDOHeader.Len));

              //mark SDO data as valid
              p_Handle_SDO_Write^.us_Status := SAFETY_SDO_DATA_VALID;

              if ( pISafety^.udVersion >= 16#1001 ) then
                SAFETY_iPushSafetyTask();
              end_if;

            elsif (UnsafeReadTransNr >= ReadFramesNeeded) then
              // We have finished all read data, go on with the next step
              UnsafeScheduler := UnsafeSchedulerDiagState;
              LastUnsafeUpdate := ops.tAbsolute;
              UnsafeReadTransNr := 0;
            else
              // time until read is not yet over - go on
              UnsafeScheduler := UnsafeSchedulerDiagState;
            end_if;
          else
            UnsafeScheduler   := UnsafeSchedulerDiagState;
          end_if;

       (* ***************************************** *)
          UnsafeSchedulerDiagState:
       (* ***************************************** *)
          // get the diag state (on user demand)
          if DiagVars.UserWantsDiagState then

            // get state via SDO communication
            SDORequestBuffer.StdHeader.CRC  := 0;                                                   // CRC is always 0 in Std communication
            SDORequestBuffer.StdHeader.Cmd  := SDO_COMMAND_GET_STATE;                               // get-state command
            SDORequestBuffer.StdHeader.Typ  := FRM_TYPECODE_STD;                                    // standard frame type
            SDORequestBuffer.StdHeader.SeqNr:= StandardSeqNr OR 16#80;                              // sequence number
            SDORequestBuffer.StdHeader.Len  := 4;                                                   // header
            SDORequestBuffer.ud_Address     := 0;
            SDORequestBuffer.us_Length      := 0;

            LastRequest := _DiagState;

#ifdef SAFETY_PROTOCOL_ANALYZER_ACTIVATED
  RecordFrame((#SDORequestBuffer)$^DINT, 1);
#endif

            //copy SDO into write-buffer
            To_StdLib.MemCpy(dest := #p_Handle_SDO_Write^.SDOStructure, source := #SDORequestBuffer, size := (sizeof(SDOHeader.StdHeader.CRC) + SDORequestBuffer.StdHeader.Len));

            //mark SDO data as valid
            p_Handle_SDO_Write^.us_Status := SAFETY_SDO_DATA_VALID;

            if ( pISafety^.udVersion >= 16#1001 ) then
              SAFETY_iPushSafetyTask();
            end_if;
          else
            UnsafeScheduler := UnsafeSchedulerDiagInfo;
          end_if;

       (* ***************************************** *)
          UnsafeSchedulerDiagInfo:
       (* ***************************************** *)

          // get the diag info (on user demand)
          if DiagVars.UserWantsDiagInfo then

            // get state via SDO communication
            StandardRequest.SDOHeader.CRC   := 0;                                                   // CRC is always 0 in Std communication
            StandardRequest.SDOHeader.Cmd   := SDO_COMMAND_GET_DIAG_INFO;                           // read command
            StandardRequest.SDOHeader.Typ   := FRM_TYPECODE_STD;                                    // standard frame type
            StandardRequest.SDOHeader.SeqNr := StandardSeqNr OR 16#80;                              // sequence number
            StandardRequest.SDOHeader.Len   := 4 + 1;                                               // header + µC-selection
            StandardRequest.aData[0]        := DiagVars.ucChoiceDiagInfo;

            LastRequest := _DiagInfo;

#ifdef SAFETY_PROTOCOL_ANALYZER_ACTIVATED
  RecordFrame((#StandardRequest)$^DINT, 1);
#endif

            //copy SDO into write-buffer
            To_StdLib.MemCpy(dest := #p_Handle_SDO_Write^.SDOStructure, source := #StandardRequest, size := (sizeof(SDOHeader.StdHeader.CRC) + StandardRequest.SDOHeader.Len));

            //mark SDO data as valid
            p_Handle_SDO_Write^.us_Status := SAFETY_SDO_DATA_VALID;

            if ( pISafety^.udVersion >= 16#1001 ) then
              SAFETY_iPushSafetyTask();
            end_if;

          else
            UnsafeScheduler := UnsafeSchedulerChannelError;
          end_if;

       (* ***************************************** *)
          UnsafeSchedulerChannelError:
       (* ***************************************** *)

          if DiagVars.UserWantsErrorInfo  then
            SDORequestBuffer.StdHeader.CRC  := 0;                                                      // CRC is always 0 in Std communication
            SDORequestBuffer.StdHeader.Cmd  := SDO_COMMAND_READ;                                       // read command
            SDORequestBuffer.StdHeader.Typ  := SDO_STD;                                                // standard frame type
            SDORequestBuffer.StdHeader.SeqNr:= StandardSeqNr OR 16#80;                                 // sequence number
            SDORequestBuffer.StdHeader.Len  := 4 + 4 + 1;                                              // header + destination address + length of data
            SDORequestBuffer.ud_Address     := SDO_ADDRESS_ERROR_MEM;                                  // address of error memory
            SDORequestBuffer.us_Length      := SDO_LENGTH_ERROR_MESSAGE;                               // length of data (first byte contains number of following values + number of channels)
            if remainingPacketlength <> 0 then
              // set offset if more than one package
              SDORequestBuffer.ud_Address     := (SDO_ADDRESS_ERROR_MEM + actoffset);                  // address of error memory
              // set new length for next package
              if remainingPacketlength > SDO_LENGTH_ERROR_MESSAGE then
                SDORequestBuffer.us_Length      := SDO_LENGTH_ERROR_MESSAGE;
              else
                SDORequestBuffer.us_Length      := remainingPacketlength$USINT;
              end_if;
            end_if;

            LastRequest := _ErrorChannelInfo;

#ifdef SAFETY_PROTOCOL_ANALYZER_ACTIVATED
  RecordFrame((#StandardRequest)$^DINT, 1);
#endif

            //copy SDO into write-buffer
            To_StdLib.MemCpy(dest := #p_Handle_SDO_Write^.SDOStructure, source := #SDORequestBuffer, size := (sizeof(SDOHeader.StdHeader.CRC) +  SDORequestBuffer.StdHeader.Len));

            //mark SDO data as valid
            p_Handle_SDO_Write^.us_Status := SAFETY_SDO_DATA_VALID;

            if ( pISafety^.udVersion >= 16#1001 ) then
              SAFETY_iPushSafetyTask();
            end_if;

          else
            UnsafeScheduler := UnsafeSchedulerGetDiagVars;
          end_if;

        else
          if bd_LogOnceMarker.InvalidSchedulerState = FALSE then
            bd_LogOnceMarker.InvalidSchedulerState := TRUE;
            bd_AlreadyLoggedMarker.InvalidSchedulerState := TRUE;
            LogError("@ZZZZ (SafetyCDIAS_Base::UpdateCy) [SL] Undefined Scheduler-State");
          end_if;
        end_case;

      end_while;
    end_if;
  end_if;

  // at the first run we write all variables independent of any changes
  if RunState > OldRunState then
    SendAllUnsafeValues();
  end_if;
  OldRunState := RunState;

//============================ Profiler start======================================================
#ifdef  DM_Profiler
  StopTimeMeasurement(usMode := DMTIME_CY);
#endif
//============================ Profiler end========================================================

END_FUNCTION

FUNCTION VIRTUAL GLOBAL SafetyCDIAS_Base::GetModuleType
	VAR_OUTPUT
		ui_ModuleType 	: UINT;
	END_VAR

  ui_ModuleType := TYPE_SAFETY_MODULE;

END_FUNCTION

FUNCTION VIRTUAL SafetyCDIAS_Base::AddModuleToSafetyTask
	VAR_OUTPUT
		sd_retval 	: DINT;
	END_VAR

  //register module as safety module in OS and receive pointers on SDO buffers
  sd_retval := SAFETY_iAddModuleToSafetyTask( uiMaster  := 0
                                            , pucNode   := p_ObjectPath
                                            , pucRdSDO  := ( #p_Handle_SDO_Read )$^UDINT
                                            , pucWrSDO  := ( #p_Handle_SDO_Write )$^UDINT
                                            );

  //look for an error
	if ( sd_retval ) then
    State.uiIO_Flags				          := 0;
		State.uiIO_Flags.NoCalibration	  := 1;
		State.uiIO_Flags.PhysicAccessOff  := 1;

    LogError("@ZZZZ (SafetyCDIAS_Base::AddModuleToSafetyTask) Module not added to Safety Communication Task");
